Staubli VAL3: loadPROG.pgx

public program loadPROG(num x_nLib, num& x_nResult)
  local string l_sPath
  local num l_nClock
begin
  l_nClock=clock()
  if x_nLib>=0

    l_sPath="Disk://data/CustomerLib/lib"+toString("",x_nLib)+"/savePROG"
    x_nResult=progTemp:libLoad(l_sPath)
    if x_nResult!=0
      popUpMsg("1")
      call rs:setAlarm(300,0)
    endIf
  else
    call rs:setAlarm(302,0)
  endIf
  logMsg(progTemp:libPath()+",耗时:"+toString(".3",clock()-l_nClock))

end
